FUNCTION_BLOCK FB_PendantSetFocusState EXTENDS FB_PendantState
VAR_INPUT
END_VAR
VAR_OUTPUT
END_VAR
VAR
	Stage 					: UINT;
	tonCount 				: TON:= (PT:=T#1S);
	fCurrentFocusPosition 	: LREAL;
	fSmallStep				: LREAL := 0.1;
	fBigStep				: LREAL := 1.0;
	fSetFocusPosition		: LREAL;
	sSetFocusPosition		: STRING;
	nFocusRightLength 		: UINT;
	
	bBlockChange			: BOOL := FALSE;
	bToIdle					: BOOL := FALSE;
	//Hex stuff
	aTxHexData				: ARRAY[0..2] OF BYTE;
	tonDelay				: TON:= (PT:=T#20MS);
END_VAR

METHOD FoundError : BOOL
Stage := 0;
tonDelay(IN:=FALSE);
tonCount(IN:=FALSE);
pPendant^.SetState(pPendant^.fbPendantErrorState);
END_METHOD

METHOD RunState : BOOL
CASE Stage OF
	0:
		fCurrentFocusPosition := F_RoundLREAL(pPendant^.ipFocus.Position,3);
		IF pPendant^._FastMove THEN
			IF pPendant^._MovePositive THEN
				fSetFocusPosition := fCurrentFocusPosition + fBigStep;
			ELSE
				fSetFocusPosition := fCurrentFocusPosition - fBigStep;
			END_IF
		ELSE
			IF pPendant^._MovePositive THEN
				fSetFocusPosition := fCurrentFocusPosition + fSmallStep;
			ELSE
				fSetFocusPosition := fCurrentFocusPosition - fSmallStep;
			END_IF
		END_IF
		pPendant^.ipFocus.Position := fSetFocusPosition;
		Stage := Stage +1;
	1:
		// Block State Change while full text is send -> to not run into issues with commands
		// Does not include Error State
		bBlockChange := TRUE;
		IF NOT pPendant^.fbSendHex.Busy OR pPendant^.fbSendString.Busy THEN
			Stage := Stage +1;
		END_IF
	2: 
		// send sequence for two line text. For first line: fe, 01, 00, 0c, first 8 char, second 8 char
		HEXSTR_TO_DATA('fe', ADR(aTxHexData), SIZEOF(aTxHexData));
		pPendant^.fbSendHex(
				pSendData:= ADR(aTxHexData),
				Length	:= 1,
				TXbuffer:= TxBufferPendant,
				Busy=>,
				Error=> );
		IF NOT pPendant^.fbSendHex.Busy THEN
			Stage := Stage +1;
		END_IF
	3: 
		HEXSTR_TO_DATA('01', ADR(aTxHexData), SIZEOF(aTxHexData));
		pPendant^.fbSendHex(
				pSendData:= ADR(aTxHexData),
				Length	:= 1,
				TXbuffer:= TxBufferPendant,
				Busy=>,
				Error=> );
		IF NOT pPendant^.fbSendHex.Busy THEN
			Stage := Stage +1;
		END_IF
	4: 
		HEXSTR_TO_DATA('00', ADR(aTxHexData), SIZEOF(aTxHexData));
		pPendant^.fbSendHex(
				pSendData:= ADR(aTxHexData),
				Length	:= 1,
				TXbuffer:= TxBufferPendant,
				Busy=>,
				Error=> );
		IF NOT pPendant^.fbSendHex.Busy THEN
			Stage := Stage +1;
		END_IF
	5:	
		HEXSTR_TO_DATA('0c', ADR(aTxHexData), SIZEOF(aTxHexData));
		pPendant^.fbSendHex(
				pSendData:= ADR(aTxHexData),
				Length	:= 1,
				TXbuffer:= TxBufferPendant,
				Busy=>,
				Error=> );
		IF NOT pPendant^.fbSendHex.Busy THEN
			Stage := Stage +1;
		END_IF
	6:
		// send first 8 characters
		pPendant^.fbSendString(SendString:= 'Focus 1-',
					TXbuffer:= TxBufferPendant,
					Busy=>,
					Error=> );
		IF NOT pPendant^.fbSendString.Busy  THEN
			Stage := Stage +1;
		END_IF
	7: 
		tonDelay(IN:=TRUE);
		IF tonDelay.Q THEN
			tonDelay(IN:=FALSE);
			Stage:=Stage +1;
		END_IF
	8:
		// send second characters (8 max)
		pPendant^.fbSendString(SendString:= '17mm    ',
					TXbuffer:= TxBufferPendant,
					Busy=>,
					Error=> );
		IF NOT pPendant^.fbSendString.Busy  THEN
			Stage := Stage +1;
		END_IF
	9: 
		tonDelay(IN:=TRUE);
		IF tonDelay.Q THEN
			tonDelay(IN:=FALSE);
			Stage:=Stage +1;
		END_IF
	10: 
		// second line: fe, c0, 00, 0b, first 8 char, second 8 char
		HEXSTR_TO_DATA('fe', ADR(aTxHexData), SIZEOF(aTxHexData));
		pPendant^.fbSendHex(
				pSendData:= ADR(aTxHexData),
				Length	:= 1,
				TXbuffer:= TxBufferPendant,
				Busy=>,
				Error=> );
		IF NOT pPendant^.fbSendHex.Busy THEN
			Stage := Stage +1;
		END_IF
	11: 
		HEXSTR_TO_DATA('c0', ADR(aTxHexData), SIZEOF(aTxHexData));
		pPendant^.fbSendHex(
				pSendData:= ADR(aTxHexData),
				Length	:= 1,
				TXbuffer:= TxBufferPendant,
				Busy=>,
				Error=> );
		IF NOT pPendant^.fbSendHex.Busy THEN
			Stage := Stage +1;
		END_IF
	12: 
		HEXSTR_TO_DATA('00', ADR(aTxHexData), SIZEOF(aTxHexData));
		pPendant^.fbSendHex(
				pSendData:= ADR(aTxHexData),
				Length	:= 1,
				TXbuffer:= TxBufferPendant,
				Busy=>,
				Error=> );
		IF NOT pPendant^.fbSendHex.Busy THEN
			Stage := Stage +1;
		END_IF
	13:	
		HEXSTR_TO_DATA('0b', ADR(aTxHexData), SIZEOF(aTxHexData));
		pPendant^.fbSendHex(
				pSendData:= ADR(aTxHexData),
				Length	:= 1,
				TXbuffer:= TxBufferPendant,
				Busy=>,
				Error=> );
		IF NOT pPendant^.fbSendHex.Busy THEN
			Stage := Stage +1;
		END_IF
	14:
		sSetFocusPosition := CONCAT(LREAL_TO_STRING(fSetFocusPosition),'        ');
		// send first 8 characters
		pPendant^.fbSendString(SendString:= MID(sSetFocusPosition,8,1),
					TXbuffer:= TxBufferPendant,
					Busy=>,
					Error=> );
		IF NOT pPendant^.fbSendString.Busy  THEN
			Stage := Stage +1;
		END_IF
	15: 
		tonDelay(IN:=TRUE);
		IF tonDelay.Q THEN
			tonDelay(IN:=FALSE);
			Stage:=Stage +1;
		END_IF
	16:
		pPendant^.fbSendString(SendString:= 'mm      ',
					TXbuffer:= TxBufferPendant,
					Busy=>,
					Error=> );
		IF NOT pPendant^.fbSendString.Busy  THEN
			// unblock State change
			bBlockChange := FALSE;
			Stage := Stage +1;
		END_IF
	17:
		tonCount(IN:=TRUE);
		IF tonCount.Q THEN
			tonCount(IN:=FALSE);
			//restart
			Stage:=0;
		END_IF
END_CASE

IF bToIdle THEN
	THIS^.ToIdle();
END_IF
END_METHOD

PROPERTY StateID : STRING
GET
StateID := 'Set Focus State';
END_GET
END_PROPERTY

METHOD ToIdle : BOOL
IF NOT bBlockChange THEN
	Stage := 0;
	tonDelay(IN:=FALSE);
	tonCount(IN:=FALSE);
	bToIdle := FALSE;
	pPendant^.SetState(pPendant^.fbPendantIdleState);
ELSE
	bToIdle := TRUE;
END_IF
END_METHOD

END_FUNCTION_BLOCK

(* stored: Version 1.1.0.1, ProductVersion 3.1.4024.15
   POU FB_PendantSetFocusState: Id {a4eff9c0-f8b9-4f55-9af3-e35d7167e3b3}, SpecialFunc None
   Method FoundError: Id {3e229a2b-14ec-43de-87cb-0decc0ba98b4}
   Method RunState: Id {4d5849c6-edcd-4a06-a85d-95b4e4592d6a}
   Property StateID: Id {82c35322-db03-46b5-a0d2-1deb70d03bdc}
   Get Get: Id {382729b0-d969-4bc1-bc38-e737cc38c7e2}
   Method ToIdle: Id {de27c716-97b2-47e9-ad59-25d6dee11c9f} *)
